Yaskawa INFORM job: HOMEX1000.JBI

/JOB
//NAME HOMEX1000
//POS
///NPOS 0,0,0,1,0,0
///TOOL 0
///POSTYPE BASE
///RECTAN
///RCONF 0,0,0,0,0,0,0,0
P0000=1000.000,270.000,0.000,180.00,0.00,90.00
//INST
///DATE 2026/10/14 18:15
///ATTR SC,RW
///GROUP1 RB1
NOP
MOVJ P000 VJ=25.00 PL=0
END
